(* IEC 61131-3 sources: crb-codesys/retrieval/output/codesys_repo/重型运输系统/healthydata/global, 5 files *)

(* ---- gCan.st ---- *)
{attribute 'qualified_only'}
VAR_GLOBAL
	C6TxMsg			AT%QW00		:Can_BUS_8Outputs;
	C6RxMsg			AT%IW00		:Can_BUS_8Inputs;
	C6RxCounter			 	   	:UINT;

	C3TxMsg			AT%QW52		:Can_BUS_8Outputs;
	C3RxMsg			AT%IW47		:Can_BUS_8Inputs;
	C3RxCounter			   	   	:UINT;

	C4TxMsg			AT%QW104	:Can_BUS_8Outputs;
	C4RxMsg			AT%IW94		:Can_BUS_8Inputs;
	C4RxCounter				  	:UINT;

	C2TxMsg			AT%QW156	:Can_BUS_8Outputs;
	C2RxMsg			AT%IW141	:Can_BUS_8Inputs;
	C2RxCounter			 	   	:UINT;
//(*
	C1TxMsg			AT%QW208	:Can_BUS_8Outputs;
	C1RxMsg			AT%IW188	:Can_BUS_8Inputs;
	C1RxCounter			   	   	:UINT;

	C5TxMsg			AT%QW260	:Can_BUS_8Outputs;
	C5RxMsg			AT%IW235	:Can_BUS_8Inputs;
	C5RxCounter				  	:UINT;
//*)

END_VAR

(* ---- gController.st ---- *)
{attribute 'qualified_only'}
VAR_GLOBAL
	//发送至SWMC的比例阀的控制指令
	sky		:ARRAY[0..10] OF CmdPercentSet;
	grd		:ARRAY[1..10] OF CmdPercentSet;
END_VAR

(* ---- gDev.st ---- *)
{attribute 'qualified_only'}
VAR_GLOBAL
	sky		:ARRAY[0..10] OF DeviceUnit;
	grd		:ARRAY[1..10] OF DeviceUnit;
END_VAR

(* ---- gModbus.st ---- *)
{attribute 'qualified_only'}
VAR_GLOBAL CONSTANT
	g_modbusDataSizeMax	:  UINT:=65535; // 从机保持寄存器数量
END_VAR
VAR_GLOBAL
	srv				:mdbsStruct;		//modbus-service
	modbusBuffer	:ARRAY[0..g_modbusDataSizeMax] OF WORD;	//输入寄存器数据区
END_VAR

(* ---- gUI.st ---- *)
{attribute 'qualified_only'}
VAR_GLOBAL

	mode	:UIMode;					//模式设定

	sky		:ARRAY[0..10] OF UIUnit;	//挡板2组
	grd		:ARRAY[1..10] OF UIUnit;	//挡板1组

	pid		:UiPid;						//pid测试界面参数

END_VAR
